TYPE "ST_LineStatus"
VERSION : 0.1
   STRUCT
      "LineId" : String[40];
      "Role" : DInt;
      "Owner" : String[80];
      "Revision" : UDInt;
      "LastUpdate" : LDT;
      "TimeSynchronized" : Bool;
      "Stale" : Bool;
      "SourceError" : DInt;
   END_STRUCT;
END_TYPE
